Fanuc KAREL source: kb00070.KL

-- PROVISIONAL review KL for V770-1; original PC SHA256 e391334c35fc2547b75086675e6e85d19c4da861389e1e7e917e3caee64d7785
-- Incomplete behavior may be omitted. Consult companion uncertainty JSON. Do not deploy.
PROGRAM KB00070
%NOLOCKGROUP
BEGIN
  -- UNRESOLVED_PC offsets 5-12; opcodes 9D,23
  -- UNRESOLVED_PC offsets 17-24; opcodes 9D,23
  -- UNRESOLVED_PC offsets 29-38; opcodes 3F,75
  -- UNRESOLVED_PC offsets 43-50; opcodes 9D,23
  -- UNRESOLVED_PC offsets 55-64; opcodes 3F,75
  -- UNRESOLVED_PC offsets 69-76; opcodes 9D,23
  -- UNRESOLVED_PC offsets 81-88; opcodes 9D,23
  -- UNRESOLVED_PC offsets 93-102; opcodes 3F,75
  -- UNRESOLVED_PC offsets 107-165; opcodes 27,22,22,22,2A,22,22,2A,22,22,22,2A,31
  -- UNRESOLVED_PC offsets 170-174; opcodes 7F
END KB00070
